(* ================================================================= *)
(*  ST_HandshakeBits                                                 *)
(*  通讯握手位信号结构体 - 16个Bool信号(8上游+8下游)                  *)
(*  版本: V1.1.0  日期: 2026-05-29                                    *)
(*  来源: SysLib/types/                                              *)
(* ================================================================= *)

TYPE ST_HandshakeBits :
STRUCT
    Heartbeat    : BOOL := FALSE;  // 送料心跳 - 本机翻转通知对方在线
    RequestOut   : BOOL := FALSE;  // 送料请求 - 向上游要料
    MoveBusy     : BOOL := FALSE;  // 搬运中 - 正在传输物料
    Complete     : BOOL := FALSE;  // 完成 - 传输完成确认
    Ready        : BOOL := FALSE;  // 就绪 - 设备准备好接收/发送
    Reserved1    : BOOL := FALSE;  // 预留
    Reserved2    : BOOL := FALSE;  // 预留
    Reserved3    : BOOL := FALSE;  // 预留

    RcvHeartbeat : BOOL := FALSE;  // 接料心跳 - 本机翻转通知对方在线
    RequestIn    : BOOL := FALSE;  // 进料请求 - 下游向本机要料
    DsMoveBusy   : BOOL := FALSE;  // 对方搬运中 - 下游正在接收
    DsComplete   : BOOL := FALSE;  // 对方完成 - 下游接收完成
    DsReady      : BOOL := FALSE;  // 对方就绪 - 下游设备就绪
    Reserved4    : BOOL := FALSE;  // 预留
    Reserved5    : BOOL := FALSE;  // 预留
    Reserved6    : BOOL := FALSE;  // 预留
END_STRUCT
END_TYPE
